(* IEC 61131-3 sources: plcfuzz/tools, 2 files *)

(* ---- light.st ---- *)
PROGRAM program0
  VAR
    PB1 AT %IX0.0 : BOOL;
    PB2 AT %IX0.1 : BOOL;
    LED AT %QX0.0 : BOOL;
  END_VAR

  LED := NOT(PB2) AND (LED OR PB1);
END_PROGRAM

CONFIGURATION Config0

  RESOURCE Res0 ON PLC
    TASK task0(INTERVAL := T#50ms,PRIORITY := 0);
    PROGRAM instance0 WITH task0 : program0;
  END_RESOURCE
END_CONFIGURATION

(* ---- test.il ---- *)
PROGRAM IL_TEST
VAR
    X : INT := 15;
    Z : BOOL := TRUE;
    Y : BOOL;
END_VAR

LD X
GT 10
LD Z
AND
ST Y
END_PROGRAM
